(*
SPDX-FileCopyrightText: c 2026 Oleksandr Tiutyk <trofimich@gmail.com>
SPDX-License-Identifier: MIT
License: https://opensource.org/license/mit
*)

(*!
<summary>Groups wide-string builder assignment, reuse and failure cases.</summary>
<description>
Owns the independent child instances and their fixed registration array. Use from one PLC task at a stable address.
</description>
*)

{attribute 'no_assign'}
{attribute 'no_explicit_call' := 'do not call this function block directly'}
FUNCTION_BLOCK WideStringBuilderTestGroup EXTENDS TOF_Testing.TestGroup<3>
VAR_STAT
	{attribute 'hide'}
	_ClassName : STRING := __POUNAME();
END_VAR
VAR
	_BuildEmpty : WideStringBuilderEmptyTest(name := "BuildEmpty", parent := THIS^);
	_BuildNotEmpty : WideStringBuilderContentTest(name := "BuildNotEmpty", parent := THIS^);
	_ErrorChecking : WideStringBuilderAssignmentFailureTest(name := "ErrorChecking", parent := THIS^);

	_Children : ARRAY [0.._ChildCount - 1] OF TOF_Testing.ITestElement :=
	[
		_BuildEmpty,
		_BuildNotEmpty,
		_ErrorChecking
	];
END_VAR

//! <summary>Borrows the fixed child array. Callers must not modify it.</summary>
{attribute 'monitoring' := 'call'}
PROPERTY Children : REFERENCE TO ARRAY [0.._ChildCount - 1] OF TOF_Testing.ITestElement
GET
Children REF= _Children;
END_GET
END_PROPERTY

//! <summary>Borrows the concrete class name. Callers must not modify it.</summary>
{attribute 'monitoring' := 'call'}
PROPERTY ClassName : REFERENCE TO STRING
GET
ClassName REF= _ClassName;
END_GET
END_PROPERTY

//! <summary>Borrows the compiler-initialized namespace name. Callers must not modify it.</summary>
{attribute 'monitoring' := 'call'}
PROPERTY NamespaceName : REFERENCE TO STRING
GET
NamespaceName REF= CurrentNamespace.Name;
END_GET
END_PROPERTY

//! <summary>Reports the concrete instance size in bytes.</summary>
{attribute 'monitoring' := 'call'}
PROPERTY SelfSize : ULINT
GET
SelfSize := XSIZEOF(THIS^);
END_GET
END_PROPERTY

END_FUNCTION_BLOCK

(* stored: Version 1.1.0.1
   POU WideStringBuilderTestGroup: Id {5d7007f3-aff4-4253-a0ef-a2a1e6537741}, SpecialFunc None
   Property Children: Id {2723699c-29e4-4474-9b02-ea979b878289}
   Get Get: Id {c1f87235-4185-4387-b68c-7486cb862e61}
   Property ClassName: Id {eb4dbcc0-af7c-45c8-b6d4-b447e782738e}
   Get Get: Id {63156230-677c-4847-886e-f44110132435}
   Property NamespaceName: Id {38abf450-e0e9-4b48-ad8c-23253208c2f2}
   Get Get: Id {9b8c3d0a-9464-4f14-bada-dfc420360ce1}
   Property SelfSize: Id {ea35de24-8ecc-4417-9ee2-72f99d761b43}
   Get Get: Id {bd3fcf1c-d5db-4a5e-9eeb-646484d4a16d} *)
